Fanuc KAREL source: KT00322.KL

PROGRAM KT00322
%NOLOCKGROUP
VAR
  P1: XYZWPREXT
  P2: JOINTPOS
  OUT: BOOLEAN
BEGIN
  P1.X = 1.0
  OUT = P1 <> P2
END KT00322
